(* Logix 5000 project; controller TFF vendor 1 type 14 code 107 rev 33.11; software revision 33.04; part 38 of 38 *)
(* tags used below, declared in another part *)
   Index : DINT;   // Index
   Index2 : DINT;   // Index
   Index3 : DINT;   // Index
   index4 : DINT;   // Index
   initial_distribute : FBD_BIT_FIELD_DISTRIBUTE;
   result : DINT[2];
   Temp1 : DINT;
   TIME : DINT[2];
   TimeInMicroSeconds : LINT;
   TimeInSeconds : LINT;
   TimeInSecondsDINT : DINT;
   FirstScanComplete : BOOL;   // First Scan Complete Flag
   FlowPath : FlowPath[64];   // Flow Path Array
   FlowPathControl : FlowPathControl;   // Flow Path Control
   FlowPathSetup : FlowPathSetup;   // Flow Path Setup Data
   PCV101_Control : PCV_Control;   // PCV101 Control UDT
   Phase0 : ALIAS FOR Phase[0];   // Phase 0
   SIC001 : ALIAS FOR Drive[1];
   SIC002 : ALIAS FOR Drive[2];
   SysControl : SysControl;   // General system status and command
   Valve : Valve[100];   // Valve Array
   ValveControl : ValveControl;   // Valve Control
   XV001 : ALIAS FOR Valve[0];
   XV002 : ALIAS FOR Valve[1];
   XV101 : ALIAS FOR Valve[7];
   XV102 : ALIAS FOR Valve[8];
   XV401 : ALIAS FOR Valve[9];
   XV701 : ALIAS FOR Valve[17];
   XV702 : ALIAS FOR Valve[18];
   XV704 : ALIAS FOR Valve[20];
(* Process, continued *)

ROUTINE UNIXTime   (* structured text *)
   (* ==========================================================
   	UNIXTime : Get the system time in UNIX format (Sec from 01/01/1970) in second and MicroSecond
   
   	List of treatments
   		- Get System time in MicroSecond
   		- Divide time in MicroSecond by 1000000 to get second
   		- Store time in Second
   
   -----------------------------------------------------------------------------------------------------------------------------------------------------
   	History
   		2019-DEC-24 - Merck - Q. Spindler - Initial version for Candidate Release 1.00.00.00.a
   ============================================================*)
   
   // Get System time
   GSV(WallClockTime,,CurrentValue,TIME[0]);
   
   // Store time in MicroSecond
   COP(TIME[0],TimeInMicroSeconds,1);
   
   
   // Divide time in MicroSecond by 1000000 to get second
   result[1]:=0;
   result[0]:=0;
   
   initial_distribute.Source:=TIME[1];
   initial_distribute.SourceBit:=11;
   initial_distribute.Length:=20;
   initial_distribute.DestBit:=0;
   initial_distribute.Target:=0;
   btdt(initial_distribute);
   Temp1:=initial_distribute.Dest;
   if Temp1>=1000000 then
   	result[1].11:=1;
   	Temp1:=Temp1-1000000;
   end_if;
   
   For index4:=10 to 0 by -1 do
   	Temp1:=Temp1+Temp1;
   	Temp1.0:=TIME[1].[index4];
   
   	if Temp1>=1000000 then
   		result[1].[index4]:=1;
   		Temp1:=Temp1-1000000;
   	end_if;
   End_for;
   
   For index4:=31 to 0 by -1 do
   	Temp1:=Temp1+Temp1;
   	Temp1.0:=TIME[0].[index4];
   
   	if Temp1>=1000000 then
   		result[0].[index4]:=1;
   		Temp1:=Temp1-1000000;
   	end_if;
   End_for;
   
   result[1].31:=TIME[1].31;
   
   
   // Store time in Second
   COP(result[0],TimeInSeconds,1);
   TimeInSecondsDINT := result[0];
END_ROUTINE

ROUTINE Valve   (* ladder *)
// Valve Control Routine
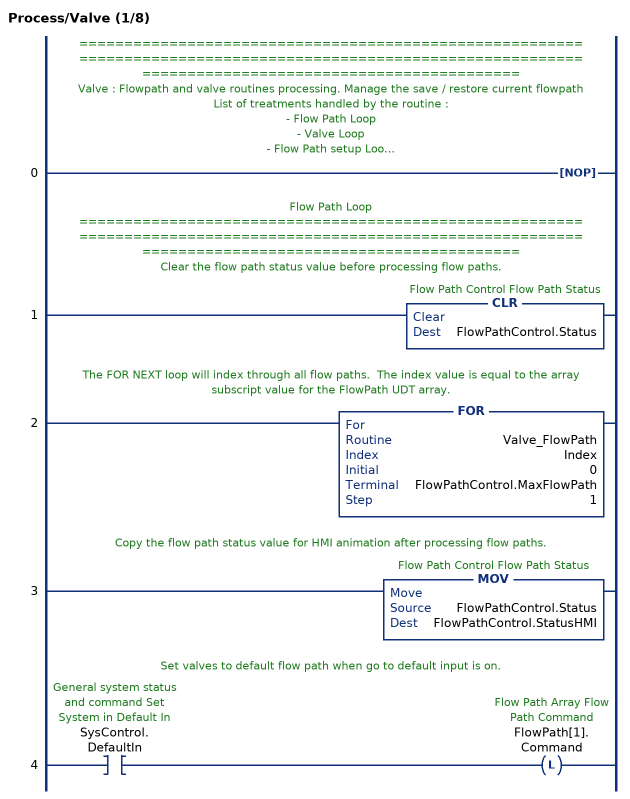
   // ==========================================================================================================================================================
   //                                                                                    Valve : Flowpath and valve routines processing. Manage the save / restore current flowpath
   //                                                     List of treatments handled by the routine :
   //                                                          - Flow Path Loop
   //                                                          - Valve Loop
   //                                                          - Flow Path setup Loop
   //                                                          - Save/restore current flowpath
   //                                                           - Valves Interlocked Status
   //                                                     -----------------------------------------------------------------------------------------------------------------------------------------------------
   //                                                     History
   // 		2019-DEC-24 - Merck - Q. Spindler - Initial version for Candidate Release 1.00.00.00.a
   //                               2020-JUN-19 - Merck - Q. Spindler - Modification for Candidate Release 1.00.00.00.c
   // - Add Valves Interlocked Status
   //                               2022-SEP-20 - Actemium - J. Jaekel - Modification for Candidate Release 1.01.00.01.a
   // - Change save flowpath logic, making it resilient from power failure when in hold
   // ========================================================================================================================================================
   0: NOP();
   // Flow Path Loop
   // ==========================================================================================================================================================
   // Clear the flow path status value before processing flow paths.
   1: CLR(FlowPathControl.Status);
   // The FOR NEXT loop will index through all flow paths.  The index value is equal to the array subscript value for the FlowPath UDT array.
   2: FOR(Valve_FlowPath,Index,0,FlowPathControl.MaxFlowPath,1);
   // Copy the flow path status value for HMI animation after processing flow paths.
   3: MOV(FlowPathControl.Status,FlowPathControl.StatusHMI);
   // Set valves to default flow path when go to default input is on.
   4: XIC(SysControl.DefaultIn)OTL(FlowPath[1].Command);
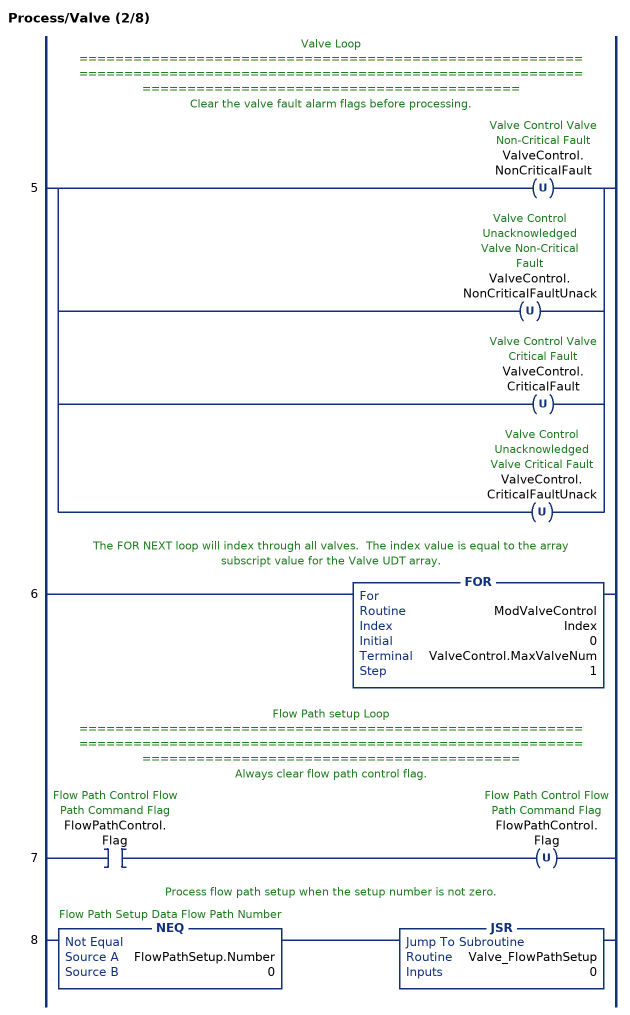
   // Valve Loop
   // ==========================================================================================================================================================
   // Clear the valve fault alarm flags before processing.
   5: [OTU(ValveControl.NonCriticalFault) ,OTU(ValveControl.NonCriticalFaultUnack) ,OTU(ValveControl.CriticalFault) ,OTU(ValveControl.CriticalFaultUnack) ];
   // The FOR NEXT loop will index through all valves.  The index value is equal to the array subscript value for the Valve UDT array.
   6: FOR(ModValveControl,Index,0,ValveControl.MaxValveNum,1);
   // Flow Path setup Loop
   // ==========================================================================================================================================================
   // Always clear flow path control flag.
   7: XIC(FlowPathControl.Flag)OTU(FlowPathControl.Flag);
   // Process flow path setup when the setup number is not zero.
   8: NEQ(FlowPathSetup.Number,0)JSR(Valve_FlowPathSetup,0);
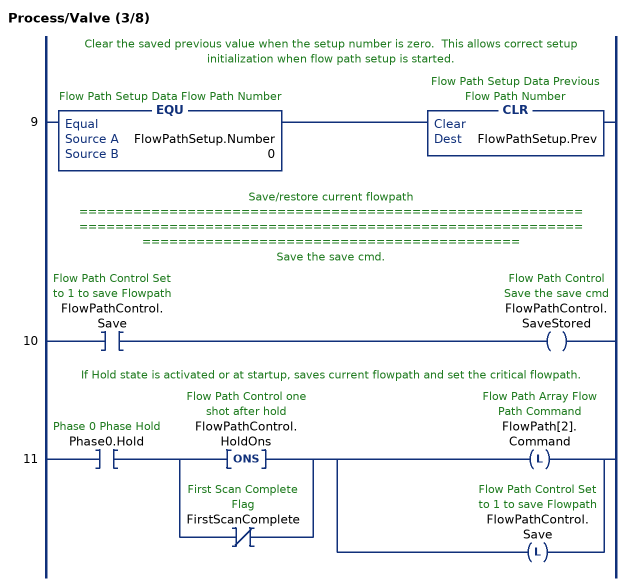
   // Clear the saved previous value when the setup number is zero.  This allows correct setup initialization when flow path setup is started.
   9: EQU(FlowPathSetup.Number,0)CLR(FlowPathSetup.Prev);
   // Save/restore current flowpath
   // ==========================================================================================================================================================
   // Save the save cmd.
   10: XIC(FlowPathControl.Save)OTE(FlowPathControl.SaveStored);
   // If Hold state is activated or at startup, saves current flowpath and set the critical flowpath.
   11: XIC(Phase0.Hold)[ONS(FlowPathControl.HoldOns) ,XIO(FirstScanComplete) ][OTL(FlowPath[2].Command) ,OTL(FlowPathControl.Save) ];
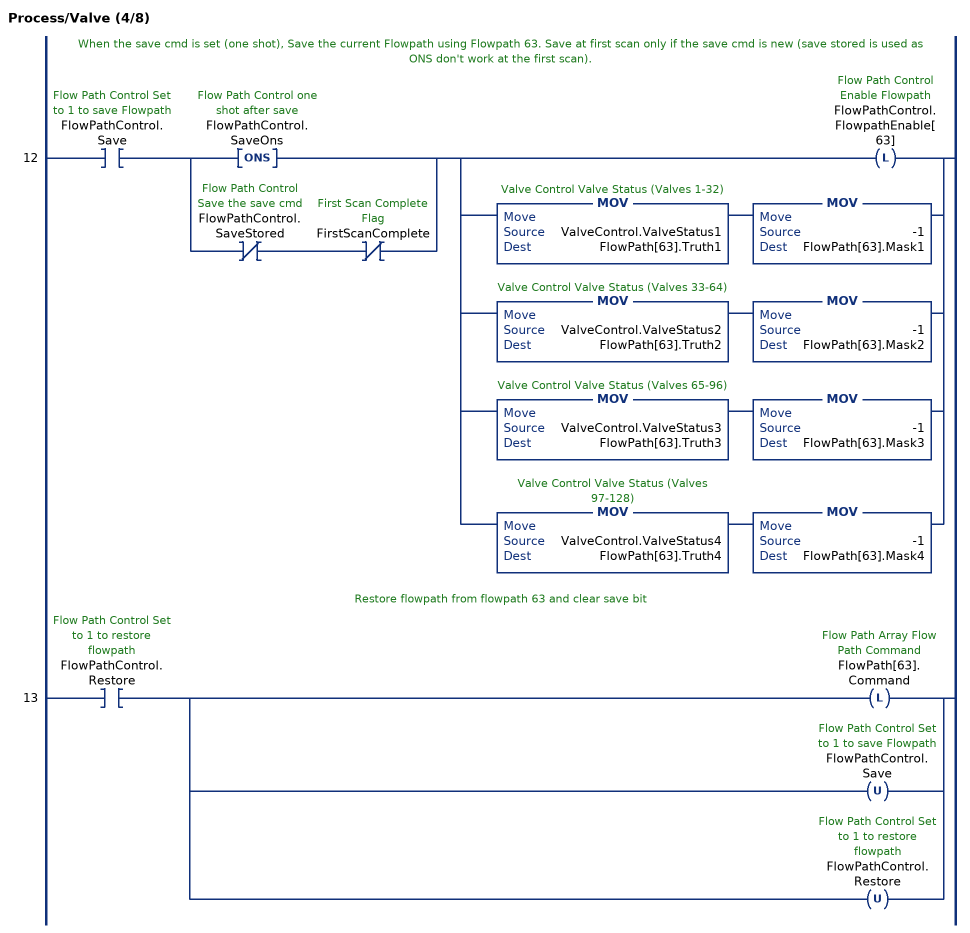
   // When the save cmd is set (one shot), Save the current Flowpath using Flowpath 63. Save at first scan only if the save cmd is new (save stored is used as ONS don't work at the first scan).
   12: XIC(FlowPathControl.Save)[ONS(FlowPathControl.SaveOns) ,XIO(FlowPathControl.SaveStored) XIO(FirstScanComplete) ][OTL(FlowPathControl.FlowpathEnable[63]) ,MOV(ValveControl.ValveStatus1,FlowPath[63].Truth1) MOV(-1,FlowPath[63].Mask1) ,MOV(ValveControl.ValveStatus2,FlowPath[63].Truth2) MOV(-1,FlowPath[63].Mask2) ,MOV(ValveControl.ValveStatus3,FlowPath[63].Truth3) MOV(-1,FlowPath[63].Mask3) ,MOV(ValveControl.ValveStatus4,FlowPath[63].Truth4) MOV(-1,FlowPath[63].Mask4) ];
   // Restore flowpath from flowpath 63 and clear save bit
   13: XIC(FlowPathControl.Restore)[OTL(FlowPath[63].Command) ,OTU(FlowPathControl.Save) ,OTU(FlowPathControl.Restore) ];
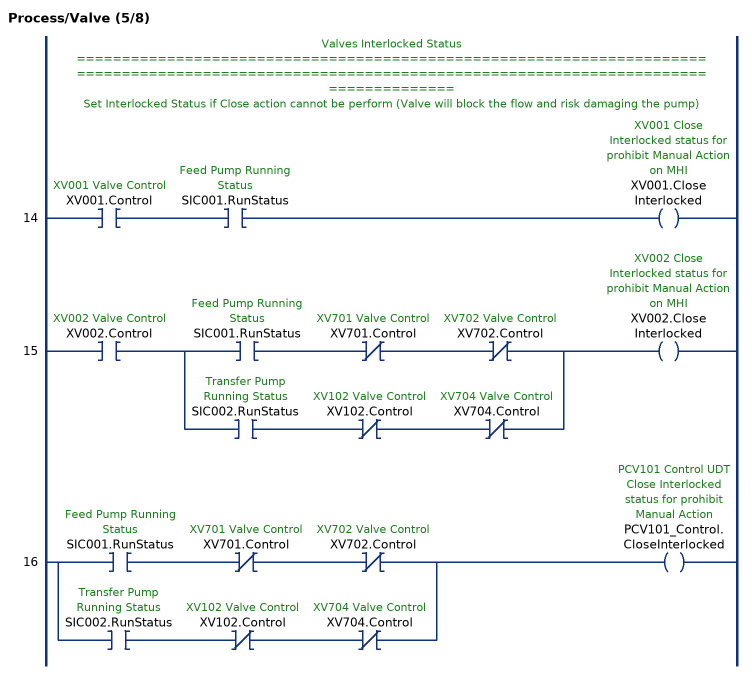
   // Valves Interlocked Status
   // ==========================================================================================================================================================
   // Set Interlocked Status if Close action cannot be perform (Valve will block the flow and risk damaging the pump)
   14: XIC(XV001.Control)XIC(SIC001.RunStatus)OTE(XV001.CloseInterlocked);
   15: XIC(XV002.Control)[XIC(SIC001.RunStatus) XIO(XV701.Control) XIO(XV702.Control) ,XIC(SIC002.RunStatus) XIO(XV102.Control) XIO(XV704.Control) ]OTE(XV002.CloseInterlocked);
   16: [XIC(SIC001.RunStatus) XIO(XV701.Control) XIO(XV702.Control) ,XIC(SIC002.RunStatus) XIO(XV102.Control) XIO(XV704.Control) ]OTE(PCV101_Control.CloseInterlocked);
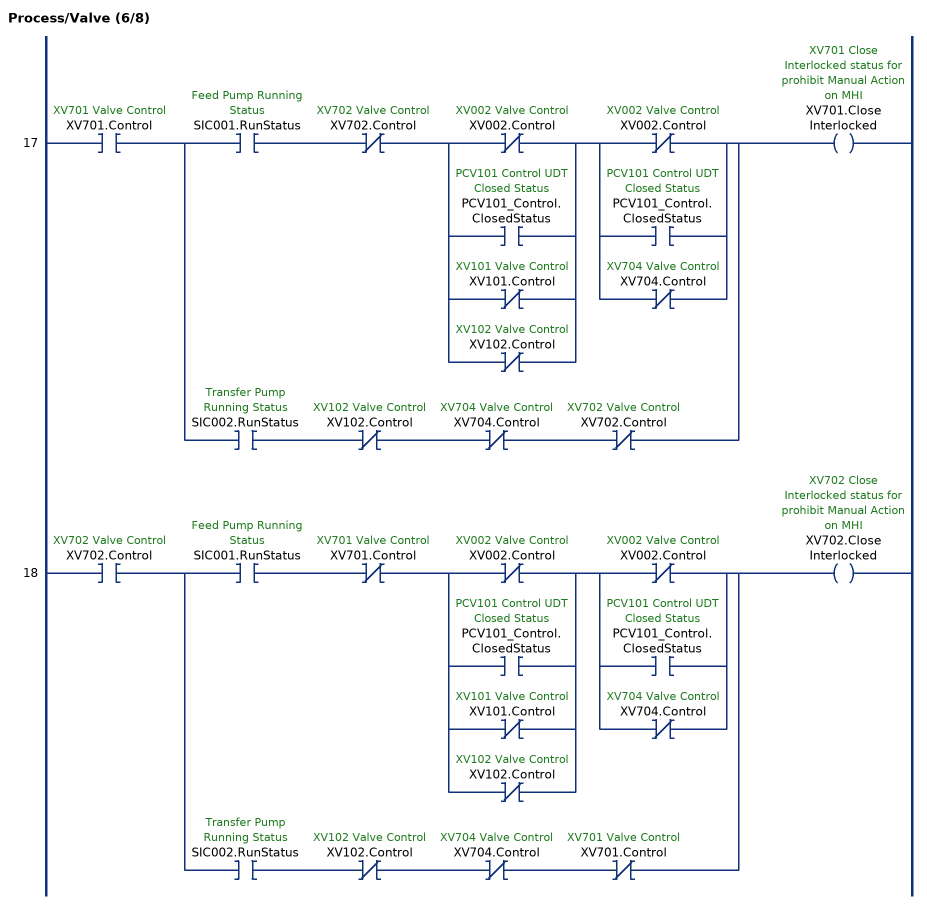
   17: XIC(XV701.Control)[XIC(SIC001.RunStatus) XIO(XV702.Control) [XIO(XV002.Control) ,XIC(PCV101_Control.ClosedStatus) ,XIO(XV101.Control) ,XIO(XV102.Control) ] [XIO(XV002.Control) ,XIC(PCV101_Control.ClosedStatus) ,XIO(XV704.Control) ] ,XIC(SIC002.RunStatus) XIO(XV102.Control) XIO(XV704.Control) XIO(XV702.Control) ]OTE(XV701.CloseInterlocked);
   18: XIC(XV702.Control)[XIC(SIC001.RunStatus) XIO(XV701.Control) [XIO(XV002.Control) ,XIC(PCV101_Control.ClosedStatus) ,XIO(XV101.Control) ,XIO(XV102.Control) ] [XIO(XV002.Control) ,XIC(PCV101_Control.ClosedStatus) ,XIO(XV704.Control) ] ,XIC(SIC002.RunStatus) XIO(XV102.Control) XIO(XV704.Control) XIO(XV701.Control) ]OTE(XV702.CloseInterlocked);
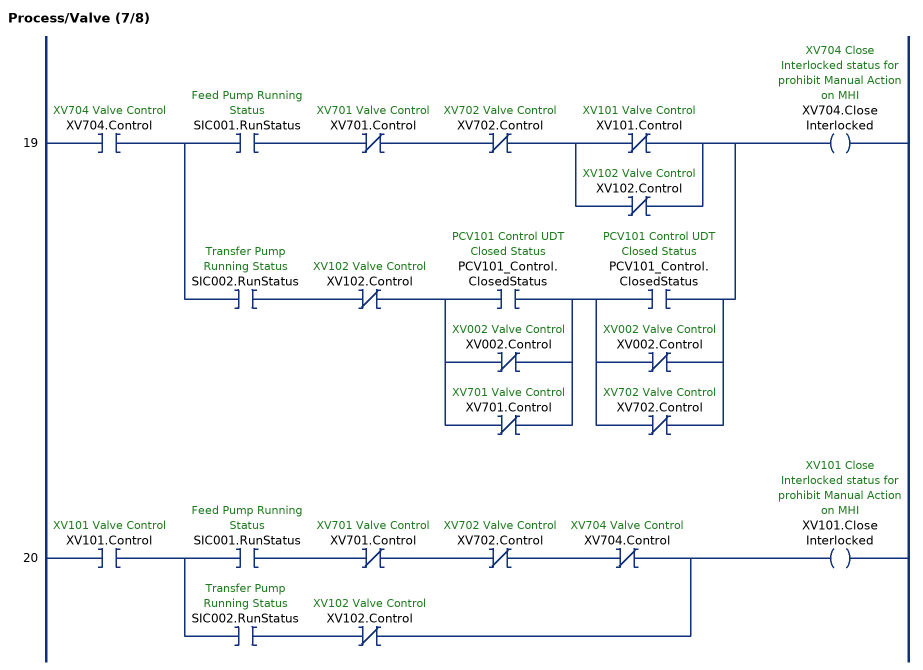
   19: XIC(XV704.Control)[XIC(SIC001.RunStatus) XIO(XV701.Control) XIO(XV702.Control) [XIO(XV101.Control) ,XIO(XV102.Control) ] ,XIC(SIC002.RunStatus) XIO(XV102.Control) [XIC(PCV101_Control.ClosedStatus) ,XIO(XV002.Control) ,XIO(XV701.Control) ] [XIC(PCV101_Control.ClosedStatus) ,XIO(XV002.Control) ,XIO(XV702.Control) ] ]OTE(XV704.CloseInterlocked);
   20: XIC(XV101.Control)[XIC(SIC001.RunStatus) XIO(XV701.Control) XIO(XV702.Control) XIO(XV704.Control) ,XIC(SIC002.RunStatus) XIO(XV102.Control) ]OTE(XV101.CloseInterlocked);
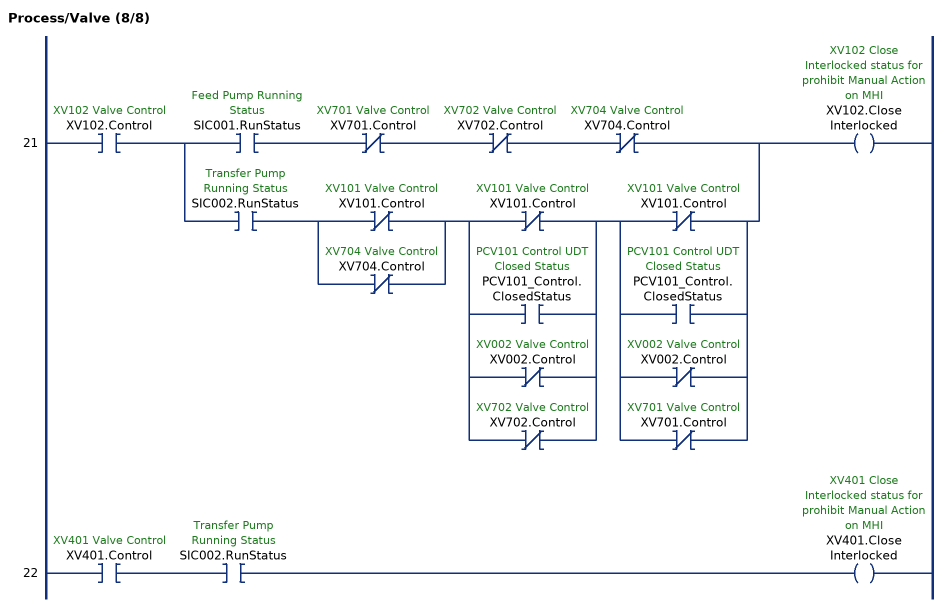
   21: XIC(XV102.Control)[XIC(SIC001.RunStatus) XIO(XV701.Control) XIO(XV702.Control) XIO(XV704.Control) ,XIC(SIC002.RunStatus) [XIO(XV101.Control) ,XIO(XV704.Control) ] [XIO(XV101.Control) ,XIC(PCV101_Control.ClosedStatus) ,XIO(XV002.Control) ,XIO(XV702.Control) ] [XIO(XV101.Control) ,XIC(PCV101_Control.ClosedStatus) ,XIO(XV002.Control) ,XIO(XV701.Control) ] ]OTE(XV102.CloseInterlocked);
   22: XIC(XV401.Control)XIC(SIC002.RunStatus)OTE(XV401.CloseInterlocked);
END_ROUTINE

ROUTINE Valve_FlowPath   (* ladder *)
// Flow Path Routine
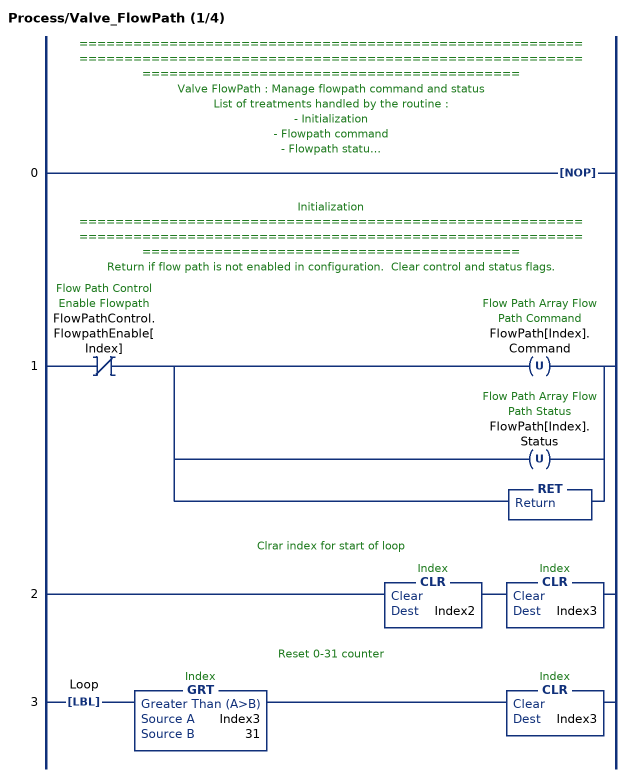
   // ==========================================================================================================================================================
   //                                                                                                  Valve FlowPath : Manage flowpath command and status
   //                                                     List of treatments handled by the routine :
   //                                                          - Initialization
   //                                                          - Flowpath command
   //                                                          - Flowpath status
   //                                                          - Reset flowpath command
   //                                                     -----------------------------------------------------------------------------------------------------------------------------------------------------
   //                                                     History
   // 		2019-DEC-24 - Merck - Q. Spindler - Initial version for Candidate Release 1.00.00.00.a
   // ========================================================================================================================================================
   0: NOP();
   // Initialization
   // ==========================================================================================================================================================
   // Return if flow path is not enabled in configuration.  Clear control and status flags.
   1: XIO(FlowPathControl.FlowpathEnable[Index])[OTU(FlowPath[Index].Command) ,OTU(FlowPath[Index].Status) ,RET() ];
   // Clrar index for start of loop
   2: CLR(Index2)CLR(Index3);
   // Reset 0-31 counter
   3: LBL(Loop)GRT(Index3,31)CLR(Index3);
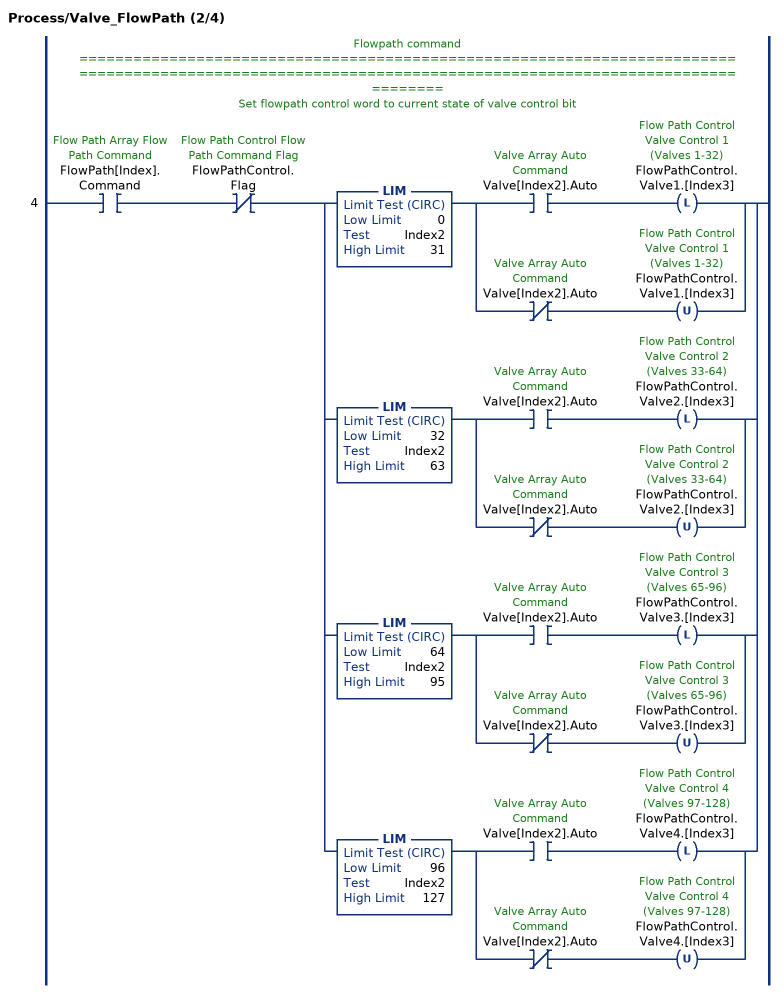
   // Flowpath command
   // ==========================================================================================================================================================
   // Set flowpath control word to current state of valve control bit
   4: XIC(FlowPath[Index].Command)XIO(FlowPathControl.Flag)[LIM(0,Index2,31) [XIC(Valve[Index2].Auto) OTL(FlowPathControl.Valve1.[Index3]) ,XIO(Valve[Index2].Auto) OTU(FlowPathControl.Valve1.[Index3]) ] ,LIM(32,Index2,63) [XIC(Valve[Index2].Auto) OTL(FlowPathControl.Valve2.[Index3]) ,XIO(Valve[Index2].Auto) OTU(FlowPathControl.Valve2.[Index3]) ] ,LIM(64,Index2,95) [XIC(Valve[Index2].Auto) OTL(FlowPathControl.Valve3.[Index3]) ,XIO(Valve[Index2].Auto) OTU(FlowPathControl.Valve3.[Index3]) ] ,LIM(96,Index2,127) [XIC(Valve[Index2].Auto) OTL(FlowPathControl.Valve4.[Index3]) ,XIO(Valve[Index2].Auto) OTU(FlowPathControl.Valve4.[Index3]) ] ];
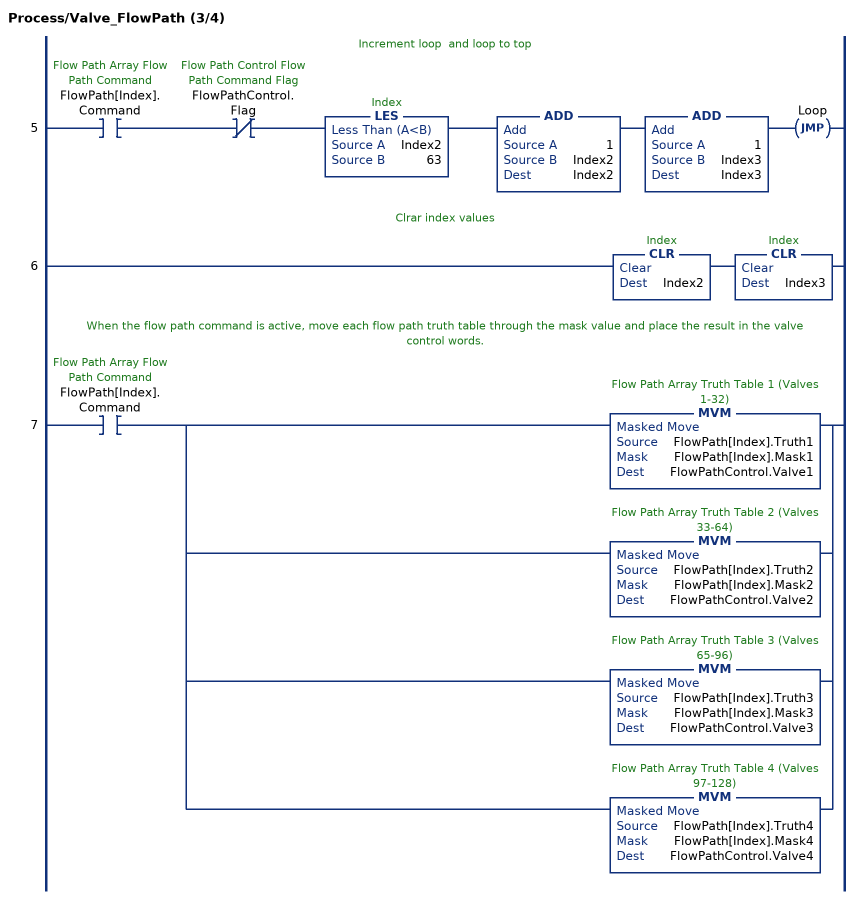
   // Increment loop  and loop to top
   5: XIC(FlowPath[Index].Command)XIO(FlowPathControl.Flag)LES(Index2,63)ADD(1,Index2,Index2)ADD(1,Index3,Index3)JMP(Loop);
   // Clrar index values
   6: CLR(Index2)CLR(Index3);
   // When the flow path command is active, move each flow path truth table through the mask value and place the result in the valve control words.
   7: XIC(FlowPath[Index].Command)[MVM(FlowPath[Index].Truth1,FlowPath[Index].Mask1,FlowPathControl.Valve1) ,MVM(FlowPath[Index].Truth2,FlowPath[Index].Mask2,FlowPathControl.Valve2) ,MVM(FlowPath[Index].Truth3,FlowPath[Index].Mask3,FlowPathControl.Valve3) ,MVM(FlowPath[Index].Truth4,FlowPath[Index].Mask4,FlowPathControl.Valve4) ];
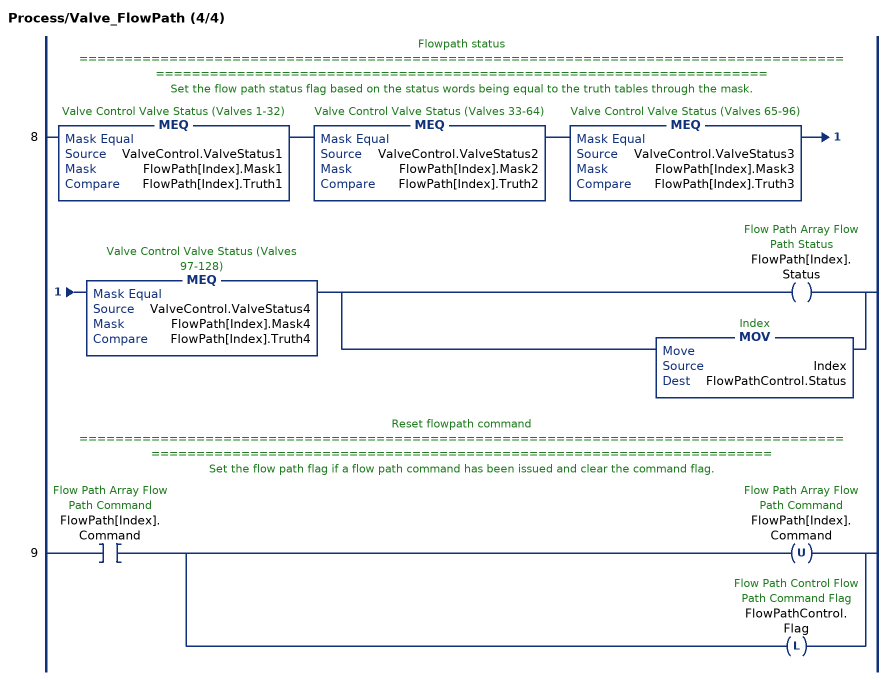
   // Flowpath status
   // =========================================================================================================================================================
   // Set the flow path status flag based on the status words being equal to the truth tables through the mask.
   8: MEQ(ValveControl.ValveStatus1,FlowPath[Index].Mask1,FlowPath[Index].Truth1)MEQ(ValveControl.ValveStatus2,FlowPath[Index].Mask2,FlowPath[Index].Truth2)MEQ(ValveControl.ValveStatus3,FlowPath[Index].Mask3,FlowPath[Index].Truth3)MEQ(ValveControl.ValveStatus4,FlowPath[Index].Mask4,FlowPath[Index].Truth4)[OTE(FlowPath[Index].Status) ,MOV(Index,FlowPathControl.Status) ];
   // Reset flowpath command
   // ==========================================================================================================================================================
   // Set the flow path flag if a flow path command has been issued and clear the command flag.
   9: XIC(FlowPath[Index].Command)[OTU(FlowPath[Index].Command) ,OTL(FlowPathControl.Flag) ];
END_ROUTINE

ROUTINE Valve_FlowPathSetup   (* ladder *)
// Flow Path Setup Routine
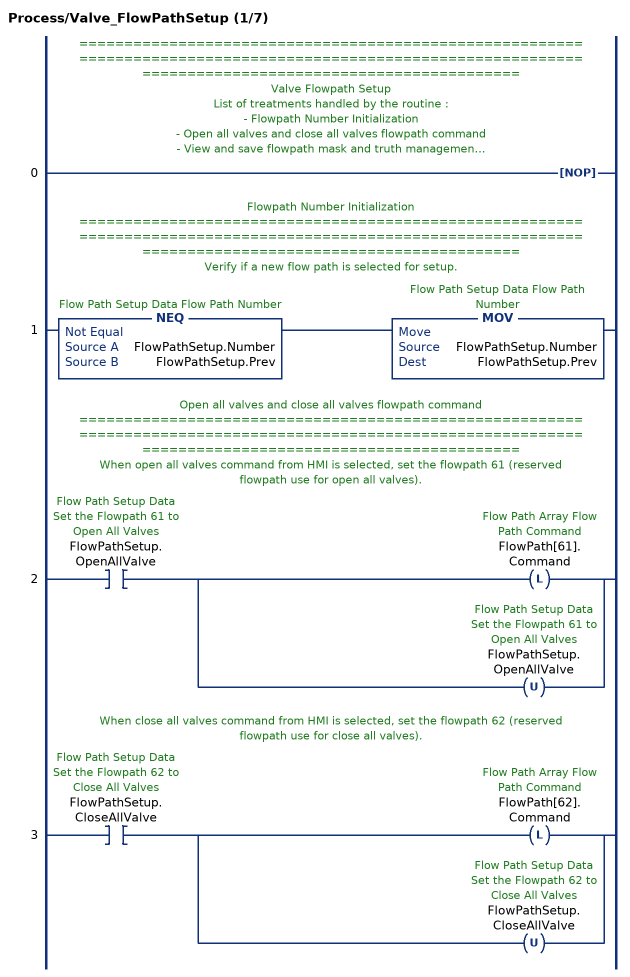
   // ==========================================================================================================================================================
   //                                                                                                                           Valve Flowpath Setup
   //                                                     List of treatments handled by the routine :
   //                                                          - Flowpath Number Initialization
   //                                                          - Open all valves and close all valves flowpath command
   //                                                          - View and save flowpath mask and truth management
   //                                                          - Apply, view mask and view truth command management
   //                                                     -----------------------------------------------------------------------------------------------------------------------------------------------------
   //                                                     History
   // 		2019-DEC-24 - Merck - Q. Spindler - Initial version for Candidate Release 1.00.00.00.a
   // ==========================================================================================================================================================
   0: NOP();
   // Flowpath Number Initialization
   // ==========================================================================================================================================================
   // Verify if a new flow path is selected for setup.
   1: NEQ(FlowPathSetup.Number,FlowPathSetup.Prev)MOV(FlowPathSetup.Number,FlowPathSetup.Prev);
   // Open all valves and close all valves flowpath command
   // ==========================================================================================================================================================
   // When open all valves command from HMI is selected, set the flowpath 61 (reserved flowpath use for open all valves).
   2: XIC(FlowPathSetup.OpenAllValve)[OTL(FlowPath[61].Command) ,OTU(FlowPathSetup.OpenAllValve) ];
   // When close all valves command from HMI is selected, set the flowpath 62 (reserved flowpath use for close all valves).
   3: XIC(FlowPathSetup.CloseAllValve)[OTL(FlowPath[62].Command) ,OTU(FlowPathSetup.CloseAllValve) ];
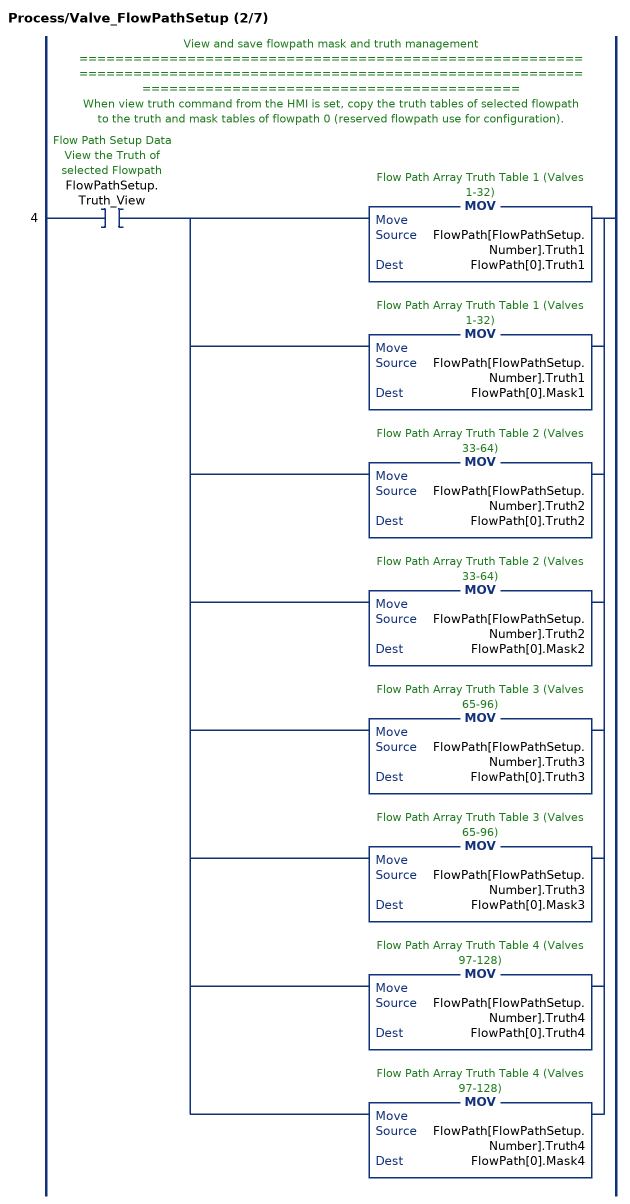
   // View and save flowpath mask and truth management
   // ==========================================================================================================================================================
   // When view truth command from the HMI is set, copy the truth tables of selected flowpath to the truth and mask tables of flowpath 0 (reserved flowpath use for configuration).
   4: XIC(FlowPathSetup.Truth_View)[MOV(FlowPath[FlowPathSetup.Number].Truth1,FlowPath[0].Truth1) ,MOV(FlowPath[FlowPathSetup.Number].Truth1,FlowPath[0].Mask1) ,MOV(FlowPath[FlowPathSetup.Number].Truth2,FlowPath[0].Truth2) ,MOV(FlowPath[FlowPathSetup.Number].Truth2,FlowPath[0].Mask2) ,MOV(FlowPath[FlowPathSetup.Number].Truth3,FlowPath[0].Truth3) ,MOV(FlowPath[FlowPathSetup.Number].Truth3,FlowPath[0].Mask3) ,MOV(FlowPath[FlowPathSetup.Number].Truth4,FlowPath[0].Truth4) ,MOV(FlowPath[FlowPathSetup.Number].Truth4,FlowPath[0].Mask4) ];
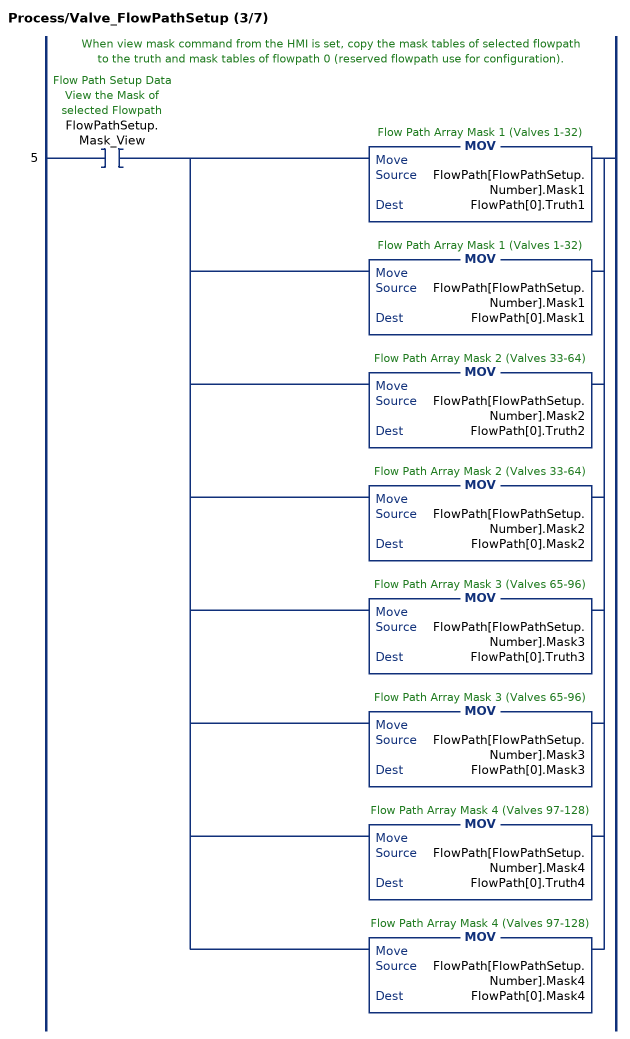
   // When view mask command from the HMI is set, copy the mask tables of selected flowpath to the truth and mask tables of flowpath 0 (reserved flowpath use for configuration).
   5: XIC(FlowPathSetup.Mask_View)[MOV(FlowPath[FlowPathSetup.Number].Mask1,FlowPath[0].Truth1) ,MOV(FlowPath[FlowPathSetup.Number].Mask1,FlowPath[0].Mask1) ,MOV(FlowPath[FlowPathSetup.Number].Mask2,FlowPath[0].Truth2) ,MOV(FlowPath[FlowPathSetup.Number].Mask2,FlowPath[0].Mask2) ,MOV(FlowPath[FlowPathSetup.Number].Mask3,FlowPath[0].Truth3) ,MOV(FlowPath[FlowPathSetup.Number].Mask3,FlowPath[0].Mask3) ,MOV(FlowPath[FlowPathSetup.Number].Mask4,FlowPath[0].Truth4) ,MOV(FlowPath[FlowPathSetup.Number].Mask4,FlowPath[0].Mask4) ];
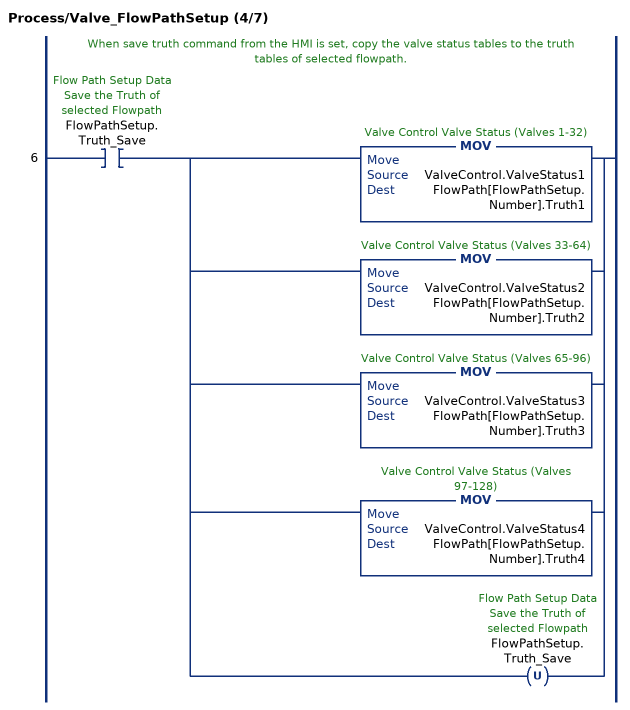
   // When save truth command from the HMI is set, copy the valve status tables to the truth tables of selected flowpath.
   6: XIC(FlowPathSetup.Truth_Save)[MOV(ValveControl.ValveStatus1,FlowPath[FlowPathSetup.Number].Truth1) ,MOV(ValveControl.ValveStatus2,FlowPath[FlowPathSetup.Number].Truth2) ,MOV(ValveControl.ValveStatus3,FlowPath[FlowPathSetup.Number].Truth3) ,MOV(ValveControl.ValveStatus4,FlowPath[FlowPathSetup.Number].Truth4) ,OTU(FlowPathSetup.Truth_Save) ];
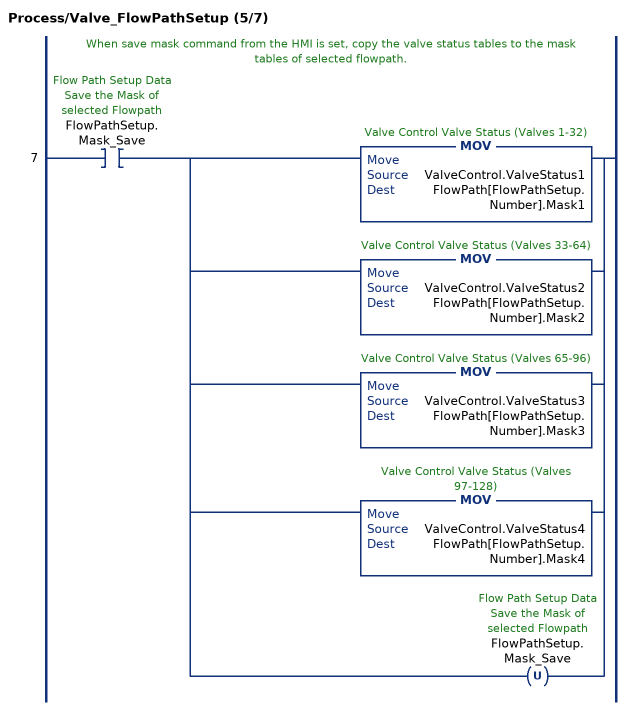
   // When save mask command from the HMI is set, copy the valve status tables to the mask tables of selected flowpath.
   7: XIC(FlowPathSetup.Mask_Save)[MOV(ValveControl.ValveStatus1,FlowPath[FlowPathSetup.Number].Mask1) ,MOV(ValveControl.ValveStatus2,FlowPath[FlowPathSetup.Number].Mask2) ,MOV(ValveControl.ValveStatus3,FlowPath[FlowPathSetup.Number].Mask3) ,MOV(ValveControl.ValveStatus4,FlowPath[FlowPathSetup.Number].Mask4) ,OTU(FlowPathSetup.Mask_Save) ];
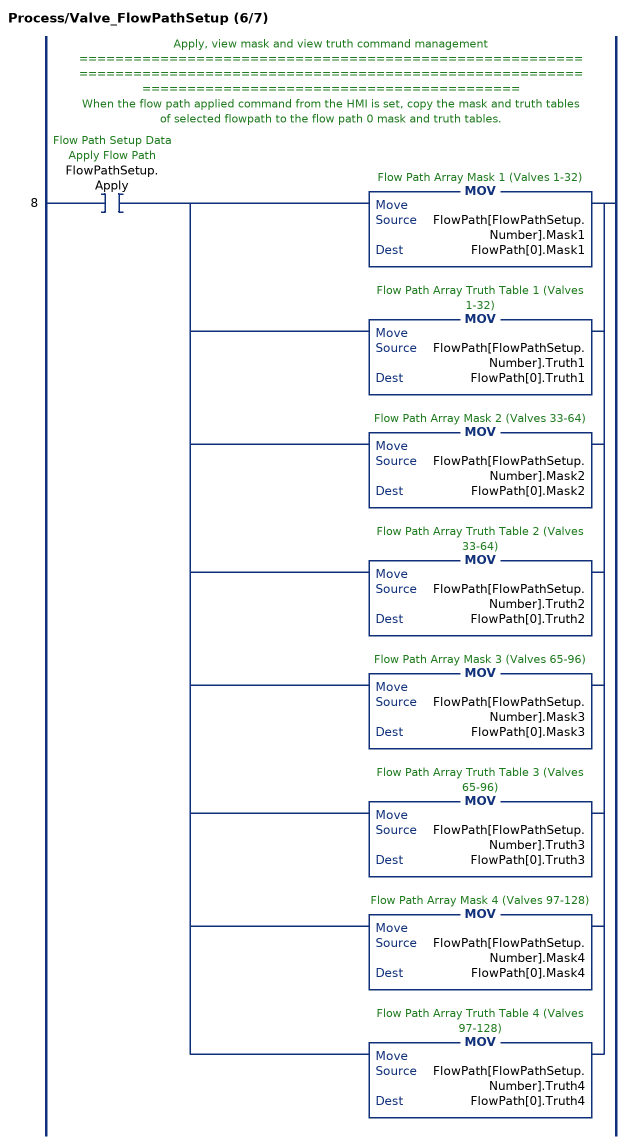
   // Apply, view mask and view truth command management
   // ==========================================================================================================================================================
   // When the flow path applied command from the HMI is set, copy the mask and truth tables of selected flowpath to the flow path 0 mask and truth tables.
   8: XIC(FlowPathSetup.Apply)[MOV(FlowPath[FlowPathSetup.Number].Mask1,FlowPath[0].Mask1) ,MOV(FlowPath[FlowPathSetup.Number].Truth1,FlowPath[0].Truth1) ,MOV(FlowPath[FlowPathSetup.Number].Mask2,FlowPath[0].Mask2) ,MOV(FlowPath[FlowPathSetup.Number].Truth2,FlowPath[0].Truth2) ,MOV(FlowPath[FlowPathSetup.Number].Mask3,FlowPath[0].Mask3) ,MOV(FlowPath[FlowPathSetup.Number].Truth3,FlowPath[0].Truth3) ,MOV(FlowPath[FlowPathSetup.Number].Mask4,FlowPath[0].Mask4) ,MOV(FlowPath[FlowPathSetup.Number].Truth4,FlowPath[0].Truth4) ];
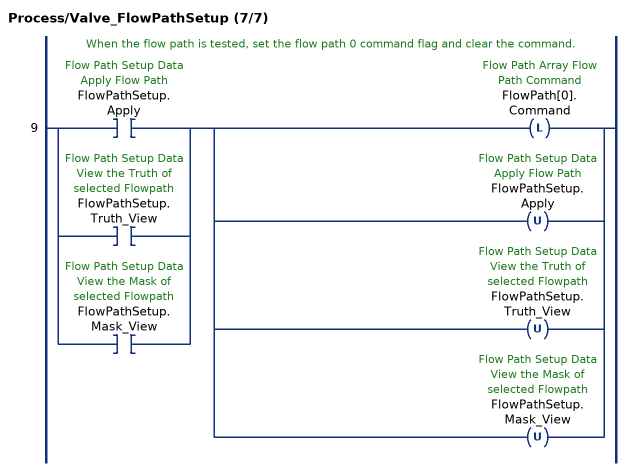
   // When the flow path is tested, set the flow path 0 command flag and clear the command.
   9: [XIC(FlowPathSetup.Apply) ,XIC(FlowPathSetup.Truth_View) ,XIC(FlowPathSetup.Mask_View) ][OTL(FlowPath[0].Command) ,OTU(FlowPathSetup.Apply) ,OTU(FlowPathSetup.Truth_View) ,OTU(FlowPathSetup.Mask_View) ];
END_ROUTINE
END_PROGRAM
